// Settable I_TelescopeStatus for tests of consumers (HMI gateway): the properties return the inputs.
FUNCTION_BLOCK FB_TelescopeStatusStub IMPLEMENTS BROTLib.I_TelescopeStatus
VAR_INPUT
	bError					: BOOL;
	nErrorID				: UDINT;
	bBusy					: BOOL;
	bIsParked				: BOOL;
	bSuspended				: BOOL;
	eLastRejectedCommand	: BROTLib.E_TCSCommand;
	eLastRejectReason		: BROTLib.E_CommandRejectReason;
	nRejectCount			: UDINT;
	fCurrentRA				: LREAL;
	fCurrentDec				: LREAL;
END_VAR

PROPERTY Error : BOOL
GET
Error := bError;
END_GET
END_PROPERTY

PROPERTY ErrorID : UDINT
GET
ErrorID := nErrorID;
END_GET
END_PROPERTY

PROPERTY Busy : BOOL
GET
Busy := bBusy;
END_GET
END_PROPERTY

PROPERTY IsParked : BOOL
GET
IsParked := bIsParked;
END_GET
END_PROPERTY

PROPERTY Suspended : BOOL
GET
Suspended := bSuspended;
END_GET
END_PROPERTY

PROPERTY LastRejectedCommand : BROTLib.E_TCSCommand
GET
LastRejectedCommand := eLastRejectedCommand;
END_GET
END_PROPERTY

PROPERTY LastRejectReason : BROTLib.E_CommandRejectReason
GET
LastRejectReason := eLastRejectReason;
END_GET
END_PROPERTY

PROPERTY RejectCount : UDINT
GET
RejectCount := nRejectCount;
END_GET
END_PROPERTY

PROPERTY CurrentRightAscension : LREAL
GET
CurrentRightAscension := fCurrentRA;
END_GET
END_PROPERTY

PROPERTY CurrentDeclination : LREAL
GET
CurrentDeclination := fCurrentDec;
END_GET
END_PROPERTY

END_FUNCTION_BLOCK

(* stored: Version 1.1.0.1, ProductVersion 3.1.4024.15
   POU FB_TelescopeStatusStub: Id {6184d763-b72f-4072-9102-f33f1a111c9a}, SpecialFunc None
   Property Error: Id {8efb484e-aeed-4917-b040-d8ff2dd81b61}
   Get Get: Id {37a7a81b-b72d-4f0b-89e2-d8b703c79ca7}
   Property ErrorID: Id {16817e2b-3b38-4095-9b98-57a3bf5dd668}
   Get Get: Id {d1afd579-b7b2-4d56-8dee-79af366293d1}
   Property Busy: Id {45b7bfd0-16d3-4793-b939-224c4490f409}
   Get Get: Id {691dc387-b576-4a39-906f-52ad738fa583}
   Property IsParked: Id {0a496587-05a1-448f-8612-733b70e2ee66}
   Get Get: Id {fcebae1c-8f8b-42ad-87de-9102ebd05829}
   Property Suspended: Id {2402739c-a84d-4852-a800-9e36ea1fc762}
   Get Get: Id {1c922f0b-0ad3-4ecf-9d4c-11de2f9d004d}
   Property LastRejectedCommand: Id {cc63b23f-415f-45bd-807c-30fb196468bd}
   Get Get: Id {267e6b69-e301-452f-b998-9562b621071f}
   Property LastRejectReason: Id {858ee852-30e6-4773-9fd2-5e8f7a77c57f}
   Get Get: Id {4f3a49f3-49b0-4b97-932d-f173ff934b5e}
   Property RejectCount: Id {ab35f529-103d-4d24-a014-f8dac5816aba}
   Get Get: Id {f0d1ca1e-ddea-40ba-ac7b-b047ed9ffad4}
   Property CurrentRightAscension: Id {e0ae9008-54f7-4696-a7f4-35322bbf57bd}
   Get Get: Id {edf0f493-784f-4af1-a299-54a4624b089f}
   Property CurrentDeclination: Id {a0cfed95-e32e-4494-b518-ccdb11311c3c}
   Get Get: Id {796b1888-5a17-4cbe-a09e-6dbf28faaa3c} *)
